{attribute 'qualified_only'}
{attribute 'strict'}
{attribute 'to_string'}
TYPE eSwitchStateType :
(
    IDLE,            // Idle - no action
    SHORT_CLICK,     // Short click
    LONG_CLICK,      // Long click
    HOLD_ON,         // Hold rising edge
	HOLD_OFF,		// Hold falling edge
    MULTI_CLICK      // Multiple click
);
END_TYPE

(* stored: Version 1.1.0.1
   DUT eSwitchStateType: Id {d36e16d9-ce68-4029-8826-9fad28d146b6} *)
